(*
SPDX-FileCopyrightText: c 2026 Oleksandr Tiutyk <trofimich@gmail.com>
SPDX-License-Identifier: MIT
License: https://opensource.org/license/mit
*)

(*!
<summary>Checks both sort directions for small strings and large DINT input.</summary>
<description>
Owns a list and its copied entries. Use from one task at a stable address.
Teardown clears surviving entries before publication.
</description>
*)

{attribute 'no_assign'}
{attribute 'no_explicit_call' := 'do not call this function block directly'}
FUNCTION_BLOCK DynamicListSortTest EXTENDS TOF_Testing.SingleCycleTest
VAR_STAT
	{attribute 'hide'}
	_ClassName : STRING := __POUNAME();
END_VAR
VAR
	_List : TOF_Collections.List<0>(valueValidator := 0);
END_VAR

(*!
<summary>Checks both sort directions for small strings and large DINT input.</summary>
*)
METHOD PROTECTED ExecuteTest
VAR
	text : ARRAY [0..15] OF STRING := [
		'S00', 'S01', 'S02', 'S03', 'S04', 'S05', 'S06', 'S07',
		'S08', 'S09', 'S10', 'S11', 'S12', 'S13', 'S14', 'S15'
	];
	i : DINT;
	value : DINT;
END_VAR
FOR i := 0 TO 15 DO
	_List.AppendCopy(value := text[i]);
END_FOR

_List.Sort(
	comparer := TOF_Comparison.StandardComparers.StringComparer,
	direction := TOF_Core.SORT_DIRECTION.DESCENDING
);

FOR i := 0 TO 15 DO
	Assert.ThatString(
		actual := _List.Get(index := i).AsString255(),
		message := TOF_Core.WideStrings.Concat255("DESCENDING STRING sort at index ", TO_WSTRING(i))
	).ToBe(expected := text[15 - i]);
END_FOR

_List.Sort(
	comparer := TOF_Comparison.StandardComparers.StringComparer,
	direction := TOF_Core.SORT_DIRECTION.ASCENDING
);

FOR i := 0 TO 15 DO
	Assert.ThatString(
		actual := _List.Get(index := i).AsString255(),
		message := TOF_Core.WideStrings.Concat255("ASCENDING STRING sort at index ", TO_WSTRING(i))
	).ToBe(expected := text[i]);
END_FOR

_List.Clear();

FOR i := 0 TO 100 DO
	value := i;
	_List.AppendCopy(value := value);
END_FOR

_List.Sort(
	comparer := TOF_Comparison.StandardComparers.DIntComparer,
	direction := TOF_Core.SORT_DIRECTION.DESCENDING
);

FOR i := 0 TO 100 DO
	Assert.ThatDInt(
		actual := _List.Get(index := i).AsDInt(),
		message := TOF_Core.WideStrings.Concat255("DESCENDING DINT sort at index ", TO_WSTRING(i))
	).ToBe(expected := 100 - i);
END_FOR

_List.Sort(
	comparer := TOF_Comparison.StandardComparers.DIntComparer,
	direction := TOF_Core.SORT_DIRECTION.ASCENDING
);

FOR i := 0 TO 100 DO
	Assert.ThatDInt(
		actual := _List.Get(index := i).AsDInt(),
		message := TOF_Core.WideStrings.Concat255("ASCENDING DINT sort at index ", TO_WSTRING(i))
	).ToBe(expected := i);
END_FOR
END_METHOD

(*!
<summary>Clears the fixture before the runner publishes the result.</summary>
<description>
Also runs after an unexpected exception interrupts the case.
</description>
*)
METHOD PROTECTED AfterTest
_List.Clear();
END_METHOD

//! <summary>Borrows the concrete class name. Callers must not modify it.</summary>
{attribute 'monitoring' := 'call'}
PROPERTY ClassName : REFERENCE TO STRING
GET
ClassName REF= _ClassName;
END_GET
END_PROPERTY

//! <summary>Borrows the compiler-initialized namespace name. Callers must not modify it.</summary>
{attribute 'monitoring' := 'call'}
PROPERTY NamespaceName : REFERENCE TO STRING
GET
NamespaceName REF= CurrentNamespace.Name;
END_GET
END_PROPERTY

//! <summary>Reports the concrete instance size in bytes.</summary>
{attribute 'monitoring' := 'call'}
PROPERTY SelfSize : ULINT
GET
SelfSize := XSIZEOF(THIS^);
END_GET
END_PROPERTY

END_FUNCTION_BLOCK

(* stored: Version 1.1.0.1
   POU DynamicListSortTest: Id {ce578c28-a57a-4bb2-9329-f95766b55d3e}, SpecialFunc None
   Method ExecuteTest: Id {7837c0e7-a25d-4bbc-a2f5-f8b88d2bc644}
   Method AfterTest: Id {2d876f56-7db8-447b-84f2-d9eb3ad84040}
   Property ClassName: Id {8de0b734-d7d1-45e5-96cc-ab4430a1bff1}
   Get Get: Id {facb1349-1cd6-4735-b2bd-fdd4d46835fa}
   Property NamespaceName: Id {87b553e1-565c-4916-af45-a4502067c245}
   Get Get: Id {0e7a2e83-7c27-4d19-96a9-31bb68bf9dd9}
   Property SelfSize: Id {183f1370-28fb-4c66-b8d4-921b7f388919}
   Get Get: Id {0547e36c-a7f5-482f-9bff-0e603d335be1} *)
